PROGRAM main
  VAR
    S1 AT %IX0.0  : BOOL; (* marcha / lote nuevo, NA *)
    S0 AT %IX0.1  : BOOL; (* parada, NC: TRUE sin pulsar *)
    B1 AT %IX0.2  : BOOL; (* sensor de piezas *)
    KM1 AT %QX0.0 : BOOL; (* motor de la cinta *)
    H1 AT %QX0.1  : BOOL; (* lote completo *)
    F_PIEZA       : R_TRIG;
    PIEZA         : BOOL; (* flanco de B1 *)
    PIEZAS        : INT; (* piezas del lote *)
    COMPLETO      : BOOL; (* lote completo *)
    F_LOTE        : R_TRIG;
    LOTE_NUEVO    : BOOL; (* flanco de COMPLETO *)
    LOTES         : INT; (* lotes completos en el turno *)
    TURNO         : BOOL; (* turno completo *)
  END_VAR
  VAR  (* added by the conversion: wires and edge detectors of the diagram *)
    _AND5_OUT : BOOL;
    _ADD9_OUT : INT;
    _SEL4_OUT : INT;
    _GE13_OUT : BOOL;
    _NOT21_OUT : BOOL;
    _AND18_OUT : BOOL;
    _SEL17_OUT : INT;
    _GE26_OUT : BOOL;
    _ADD36_OUT : INT;
    _SEL33_OUT : INT;
    _OR41_OUT : BOOL;
    _NOT45_OUT : BOOL;
    _AND40_OUT : BOOL;
  END_VAR

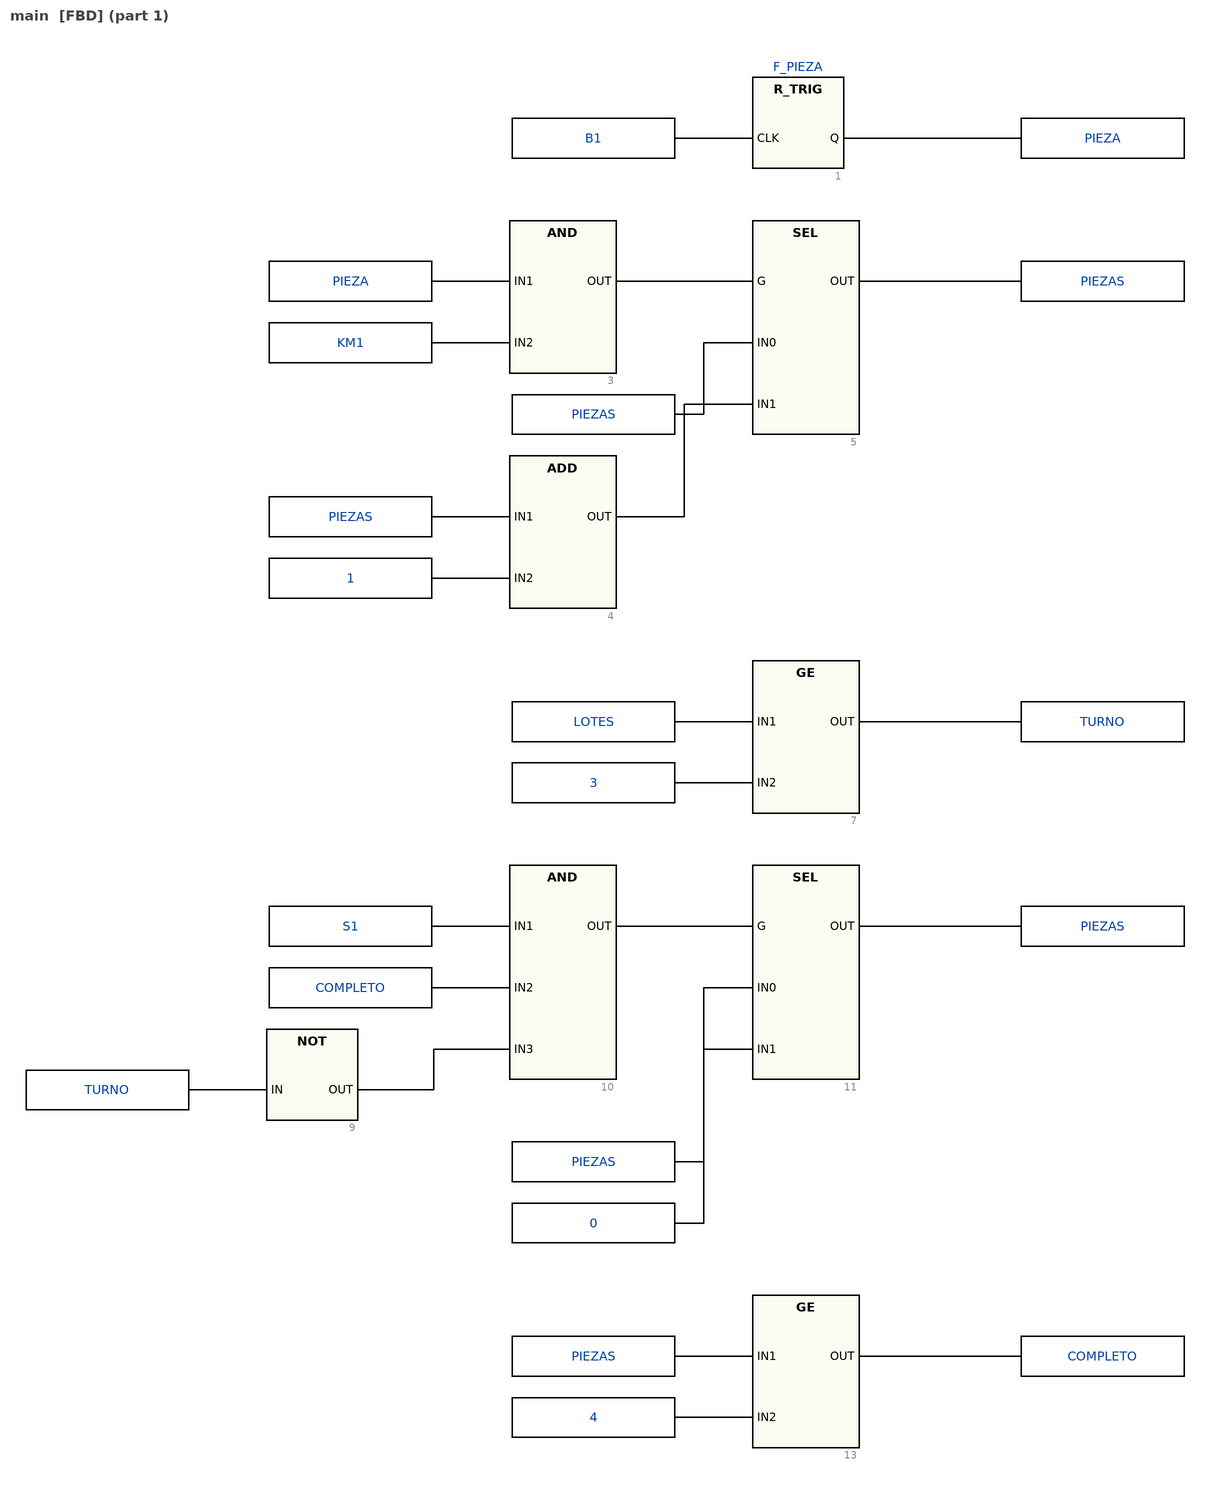
(* FBD diagram, written out as Structured Text *)
F_PIEZA(CLK := B1);
PIEZA := F_PIEZA.Q;
_AND5_OUT := PIEZA AND KM1;
_ADD9_OUT := PIEZAS + 1;
_SEL4_OUT := SEL(_AND5_OUT, PIEZAS, _ADD9_OUT);
PIEZAS := _SEL4_OUT;
_GE13_OUT := LOTES >= 3;
TURNO := _GE13_OUT;
_NOT21_OUT := NOT TURNO;
_AND18_OUT := S1 AND COMPLETO AND _NOT21_OUT;
_SEL17_OUT := SEL(_AND18_OUT, PIEZAS, 0);
PIEZAS := _SEL17_OUT;
_GE26_OUT := PIEZAS >= 4;
COMPLETO := _GE26_OUT;
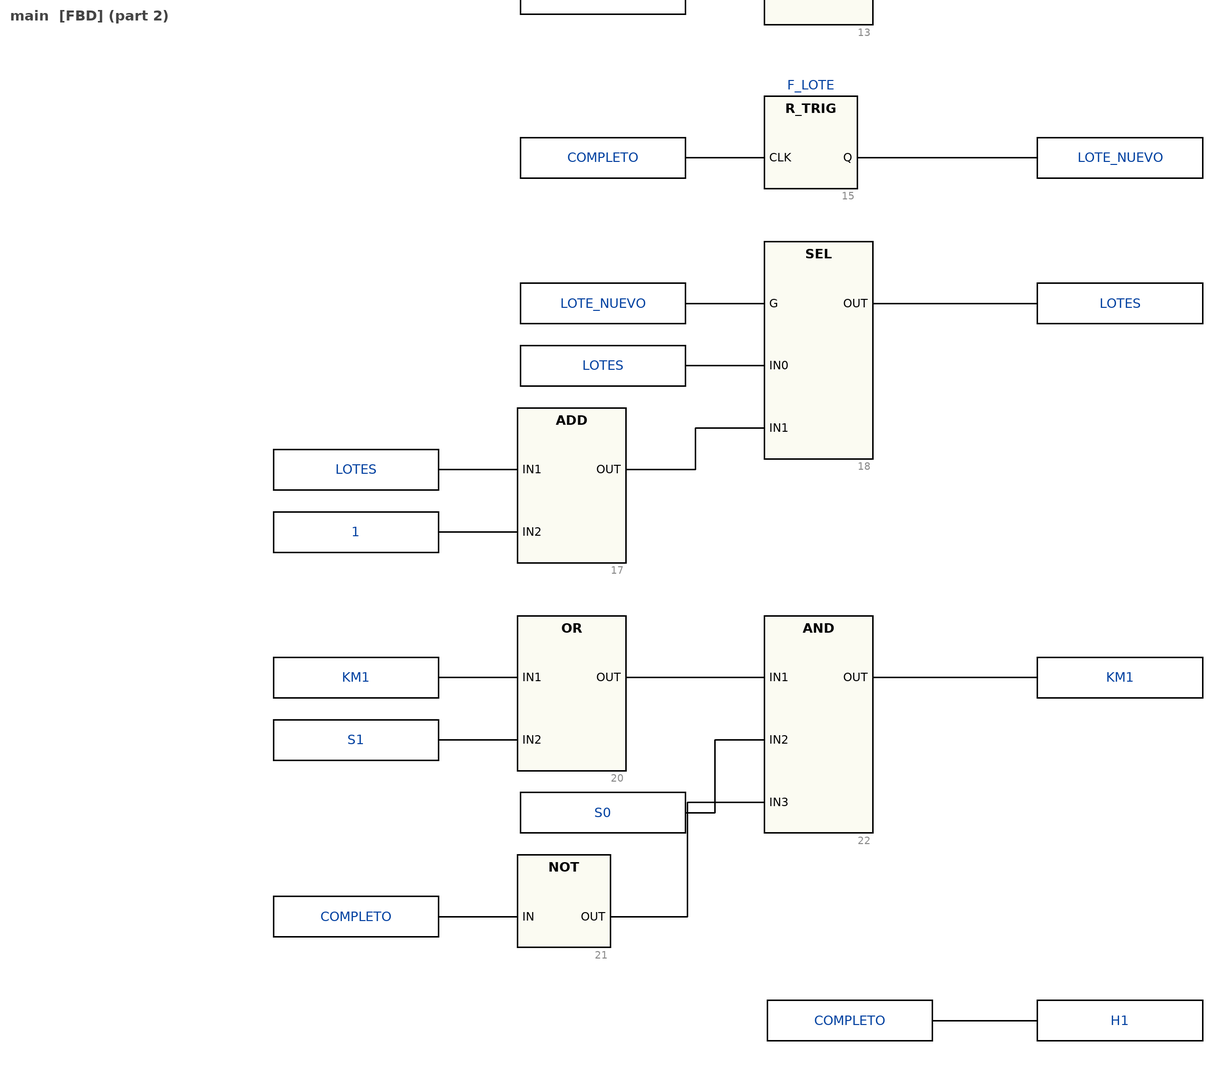
F_LOTE(CLK := COMPLETO);
LOTE_NUEVO := F_LOTE.Q;
_ADD36_OUT := LOTES + 1;
_SEL33_OUT := SEL(LOTE_NUEVO, LOTES, _ADD36_OUT);
LOTES := _SEL33_OUT;
_OR41_OUT := KM1 OR S1;
_NOT45_OUT := NOT COMPLETO;
_AND40_OUT := _OR41_OUT AND S0 AND _NOT45_OUT;
KM1 := _AND40_OUT;
H1 := COMPLETO;
END_PROGRAM
